(* IEC 61131-3 sources: trust-platform/conformance/cases/timers/cfm_timers_tp_sequence_003, 1 file *)

(* ---- program.st ---- *)
PROGRAM Main
VAR
    tp_fb : TP;
    in_tp : BOOL;
    q_tp : BOOL;
    et_tp : TIME;
END_VAR

tp_fb(IN := in_tp, PT := T#10ms, Q => q_tp, ET => et_tp);
END_PROGRAM
